{attribute 'qualified_only'}
TYPE E_FillStep :
(
	Idle,
	OpenInlet,
	Filling,
	Settle,
	Done
) UINT;
END_TYPE

(* stored: Version 1.1.0.1
   DUT E_FillStep: Id {df5fd809-eabd-4411-975d-ad3838726c88} *)
